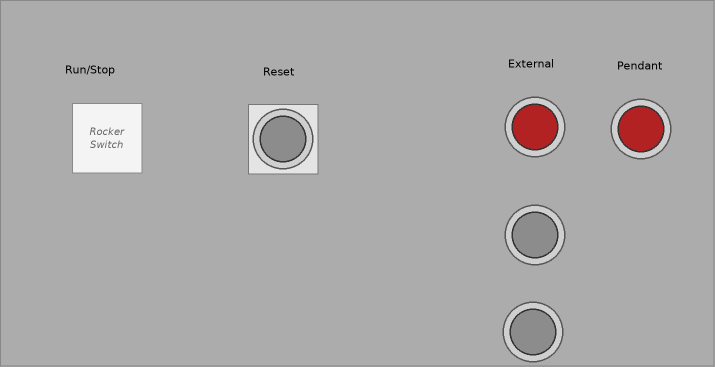
VISUALIZATION Visualization  // 715x367
    RockerSwitch (72,103 70x70), variable: bRunStop, behaviour: TOGGLE, style: Switch-RockerSwitch-Gray
    PushSwitch (248,104 70x70), variable: Estop1_RX, behaviour: TAP, style: Switch-PushSwitch-Gray
    Lamp1 (500,92 70x70), variable: not Estop1_Y, style: Lamp-Lamp1-Red
    Lamp1 (606,94 70x70), variable: not bLocalEstopFromKUKA, style: Lamp-Lamp1-Red
    Lamp1 (500,200 70x70), variable: Estop1_A, style: Lamp-Lamp1-Gray
    Lamp1 (498,297 70x70), variable: Estop1_B, style: Lamp-Lamp1-Gray
    Label (15,55 150x30), "Run/Stop"
    Label (204,57 150x30), "Reset"
    Label (456,49 150x30), "External"
    Label (565,51 150x30), "Pendant"
END_VISUALIZATION

(* stored: Version 1.1.0.1, ProductVersion 3.1.4024.12
   Visu Visualization: Id {40320f6a-8857-41e8-abc1-9a09fd87fdf0} *)
